FUNCTION FindIntField : INT
VAR_INPUT
    FieldName : STRING(254);
    JsonStr : STRING(254);
END_VAR
VAR_OUTPUT
    Valid : BOOL;
END_VAR

FindIntField := FindINTFieldFragmented(FieldName := FieldName, Str1 := JsonStr, Str2 := '', Valid => Valid);

END_FUNCTION

(* stored: Version 1.1.0.1
   POU FindIntField: Id {08b8be28-dd5e-40a3-8585-6f98ef4035d5}, SpecialFunc None *)
